FUNCTION_BLOCK BLINK
VAR_INPUT
	OnTime : TIME;
	OffTime : TIME;
END_VAR
VAR_OUTPUT
	OUT : BOOL;
END_VAR
VAR
	fbTon : TON;
	fbOff : TON;
END_VAR

fbTon.PT := OnTime;
fbOff.PT := OffTime;

fbTon.IN := NOT fbOff.Q;
fbTon();

fboff.IN := fbOff.Q;
fbOff();

OUT := fbTon.Q;

END_FUNCTION_BLOCK

(* stored: Version 1.1.0.1
   POU BLINK: Id {d9ededf5-23a2-44eb-a865-f0200f148ab1}, SpecialFunc None *)
